(* PLC project v0.5.4_.project, CODESYS CODESYS V3.5 SP19 Patch 1 *)
(* stored: creationDateTime 2026-08-04T02:31:11.4754349, modificationDateTime 2026-08-04T02:30:39.8474785 *)

PROGRAM PRG_TestSafety_LD
  VAR
    instFB_Safety_EmergencyManagement_0 : FB_Safety_EmergencyManagement;
  END_VAR

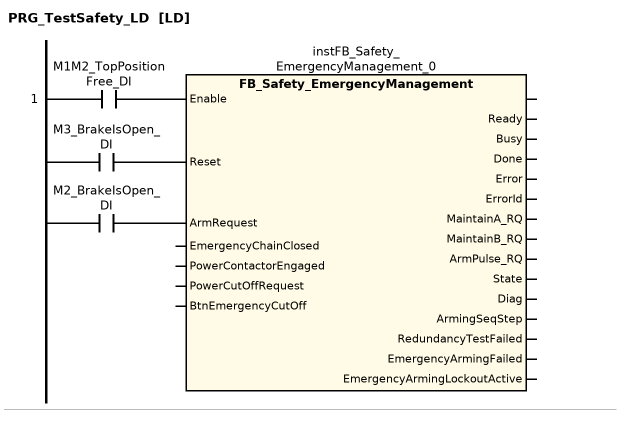
(* LD diagram, written out as Structured Text *)

instFB_Safety_EmergencyManagement_0(Enable := M1M2_TopPositionFree_DI, Reset := M3_BrakeIsOpen_DI, ArmRequest := M2_BrakeIsOpen_DI, EmergencyChainClosed := , PowerContactorEngaged := , PowerCutOffRequest := , BtnEmergencyCutOff := );
END_PROGRAM
